// TIA Portal V20 export
// export: Created 2026-10-12T05:35:23.4566716Z, ExportSetting WithDefaults, DisplayName Totally Integrated Automation Portal, DisplayVersion V20, DisplayName TIA Portal Openness, DisplayVersion V20, DisplayName TIA Portal Teamcenter Gateway, DisplayVersion V20, DisplayName TIA Portal Version Control Interface, DisplayVersion V20, DisplayName SINAMICS Startdrive Advanced, DisplayVersion V20 SP1 Update 2, DisplayName SINAMICS Startdrive G110M, G120, G120C, G120D, G120P, G115D, DisplayVersion V20 SP1 Update 2, DisplayName SINAMICS Startdrive G130, G150, S120, S150, SINAMICS MV, G220, S200, S210, DisplayVersion V20 SP1 Update 2, DisplayName STEP 7 Professional, DisplayVersion V20, DisplayName STEP 7 Safety, DisplayVersion V20, DisplayName WinCC Basic/Comfort/Advanced, DisplayVersion V20, DisplayName WinCC Professional, DisplayVersion V20, DisplayName WinCC Unified, DisplayVersion V20
FUNCTION "FRK_AlarmCapture" : Void   // FC37, SCL
{ S7_Optimized_Access := 'TRUE' }
VERSION : 0.1
// stored: AutoNumber true, IsIECCheckEnabled false, SetENOAutomatically false, UDAEnableTagReadback false
   VAR_IN_OUT
      AlarmLog : "FRK_AlarmLog";
      Core : "FRK_Core";
      Status : "ST_ModuleStatus";
   END_VAR
   VAR_TEMP
      Slot : Int;
   END_VAR
BEGIN

   #Slot := #Core.FaultSlot;
   IF #Slot < 1 OR #Slot > 16 THEN
       #Slot := 0;
   ELSIF NOT #AlarmLog.Automatic[#Slot] OR #AlarmLog.Active[#Slot].State <> 1
       OR #AlarmLog.Active[#Slot].SourcePath <> #Status.Diagnostic.SourcePath
       OR #AlarmLog.Active[#Slot].ReasonCode <> #Status.Diagnostic.ReasonCode
       OR #AlarmLog.Active[#Slot].Description <> #Status.Diagnostic.Description THEN
       #Slot := 0;
   END_IF;
   IF #Core.Exec = 3 AND NOT #Core.FaultHandled THEN
       IF #Slot = 0 THEN
           // Adopted first-outs share one active occurrence within this log.
           FOR #Slot := 1 TO 16 DO
               IF #AlarmLog.Automatic[#Slot] AND #AlarmLog.Active[#Slot].State = 1
                   AND #AlarmLog.Active[#Slot].SourcePath = #Status.Diagnostic.SourcePath
                   AND #AlarmLog.Active[#Slot].ReasonCode = #Status.Diagnostic.ReasonCode
                   AND #AlarmLog.Active[#Slot].Description = #Status.Diagnostic.Description THEN
                   EXIT;
               END_IF;
           END_FOR;
           IF #Slot > 16 THEN
               #Slot := "FRK_AlarmRaise"(AlarmLog := #AlarmLog, Diag := #Status.Diagnostic, ResetClass := 1);
           END_IF;
       END_IF;
       IF #Slot > 0 THEN
           #AlarmLog.Automatic[#Slot] := TRUE;
           #AlarmLog.Touched[#Slot] := TRUE;
       END_IF;
       #Core.FaultSlot := #Slot;
   ELSE
       #Core.FaultSlot := 0;
   END_IF;
END_FUNCTION
